(* IEC 61131-3 sources: Caravan/Archiv/12-04-19/Stations/MachineControl/MachineControl/Network/STDPLCInfoPLC, 1 file *)

(* ---- ONE_STDPLCInfoPLC_Table.st ---- *)
#define OBJECTS_CONFIG

#include <.\lsl_st_mt.h>
//Define part of class PLC_Info
#define PLC_INFO_UPDATE_TIME                    250       //Update time in cywork for CPU values
#define PLC_INFO_DEVICE_ID_CPU_REGISTER         16#0F02   //Device ID from wb_cpu_register from  FPGA
#define PLC_INFO_CPU_REGISTER_OFFSET_CPU_TEMP   16#0A     //Offset of wb_cpu_register for CPU Temperature
#define PLC_INFO_CONVERT_TO_1_10_CELSIUS        10        //Multiplier to convert temperature to 1/10°C
#include "..\..\Source\interfaces\lsl_st_pci.h"
#include "..\..\Source\interfaces\lsl_st_syssernum.h"
#include "..\..\Class\PLC_Info\XRegs.h"
#include <.\LoaderItf.h>
#include "..\..\Source\interfaces\lsl_st_sysinfo.h"

FUNCTION GLOBAL TAB ONE_STDPLCInfoPLC
-1$UINT, 0$UINT,
1$UINT, 0$UINT,

7$UDINT,
TO_UDINT(2897291062), "ASCII_BIN", 1$UINT, 20$UINT, 1$UINT,
TO_UDINT(4017734107), "GetOSVersion", 1$UINT, 2$UINT, 1$UINT,
TO_UDINT(2225119864), "MerkerEx", 1$UINT, 22$UINT, 6$UINT,
TO_UDINT(1551372421), "PLC_Info", 1$UINT, 68$UINT, 1$UINT,
TO_UDINT(1850111279), "String", 1$UINT, 10$UINT, 6$UINT,
TO_UDINT(2898603620), "StringInternal", 1$UINT, 82$UINT, 0$UINT,
TO_UDINT(3232495061), "VirtualBaseInit", 1$UINT, 3$UINT, 0$UINT,

_NO_ATTR, TO_UDINT(2882889660), "OSVERSIONPLC",

_NO_ATTR, TO_UDINT(3271492034), "GETOSVERSION_PLC",

1$UINT, TO_UDINT(884148240), "STDPLC_INFOMC1\APPLINAME\MERKEREX0",
1$UINT, TO_UDINT(2112576231), "STDPLC_INFOMC1\CPUBOARD\MERKEREX0",
1$UINT, TO_UDINT(3287353412), "STDPLC_INFOMC1\STRING0\MERKEREX0",
1$UINT, TO_UDINT(41932676), "STDPLC_INFOMC1\STRING1\MERKEREX0",
1$UINT, TO_UDINT(2235530159), "STDPLC_INFOMC1\SYSINFO\MERKEREX0",
1$UINT, TO_UDINT(3997641336), "STRINGOSVERSION_PLC\MERKEREX0",

_NO_ATTR, TO_UDINT(3849002512), "STDPLC_INFOMC1",

1$UINT, TO_UDINT(75928146), "STDPLC_INFOMC1\APPLINAME",
1$UINT, TO_UDINT(3372416669), "STDPLC_INFOMC1\CPUBOARD",
1$UINT, TO_UDINT(1828594461), "STDPLC_INFOMC1\STRING0",
1$UINT, TO_UDINT(469308299), "STDPLC_INFOMC1\STRING1",
1$UINT, TO_UDINT(882984095), "STDPLC_INFOMC1\SYSINFO",
_NO_ATTR, TO_UDINT(3965193377), "STRINGOSVERSION_PLC",

//Internal connections
0$UDINT,
11$UDINT,
TO_UDINT(8), "String0", TO_UDINT(11),
TO_UDINT(8), "String1", TO_UDINT(12),
TO_UDINT(8), "AppliName", TO_UDINT(9),
TO_UDINT(8), "CPUBoard", TO_UDINT(10),
TO_UDINT(8), "SysInfo", TO_UDINT(13),
TO_UDINT(9), "MerkerEx0", TO_UDINT(2),
TO_UDINT(10), "MerkerEx0", TO_UDINT(3),
TO_UDINT(11), "MerkerEx0", TO_UDINT(4),
TO_UDINT(12), "MerkerEx0", TO_UDINT(5),
TO_UDINT(13), "MerkerEx0", TO_UDINT(6),
TO_UDINT(14), "MerkerEx0", TO_UDINT(7),
0$UDINT,
8$UDINT,
TO_UDINT(1), "cOSVersion", TO_UDINT(14), "Data",
TO_UDINT(1), "cAsciiBin", TO_UDINT(0), "Obj_channel",
TO_UDINT(9), "DataBuffer", TO_UDINT(2), "m_udLength",
TO_UDINT(10), "DataBuffer", TO_UDINT(3), "m_udLength",
TO_UDINT(11), "DataBuffer", TO_UDINT(4), "m_udLength",
TO_UDINT(12), "DataBuffer", TO_UDINT(5), "m_udLength",
TO_UDINT(13), "DataBuffer", TO_UDINT(6), "m_udLength",
TO_UDINT(14), "DataBuffer", TO_UDINT(7), "m_udLength",

//Initialization values
0$UDINT,
10$UDINT,
TO_UDINT(2), "ThreadSafe", TO_UDINT(0),//|STDPLCInfoPLC.AppliName\STDPLC_InfoMC1\MerkerEx0.ThreadSafe;
TO_UDINT(3), "ThreadSafe", TO_UDINT(0),//|STDPLCInfoPLC.CPUBoard\STDPLC_InfoMC1\MerkerEx0.ThreadSafe;
TO_UDINT(4), "ThreadSafe", TO_UDINT(0),//|STDPLCInfoPLC.String0\STDPLC_InfoMC1\MerkerEx0.ThreadSafe;
TO_UDINT(5), "ThreadSafe", TO_UDINT(0),//|STDPLCInfoPLC.String1\STDPLC_InfoMC1\MerkerEx0.ThreadSafe;
TO_UDINT(6), "ThreadSafe", TO_UDINT(0),//|STDPLCInfoPLC.SysInfo\STDPLC_InfoMC1\MerkerEx0.ThreadSafe;
TO_UDINT(9), "SingleRealloc", TO_UDINT(1),//|STDPLCInfoPLC.STDPLC_InfoMC1\AppliName.SingleRealloc;
TO_UDINT(10), "SingleRealloc", TO_UDINT(1),//|STDPLCInfoPLC.STDPLC_InfoMC1\CPUBoard.SingleRealloc;
TO_UDINT(11), "SingleRealloc", TO_UDINT(1),//|STDPLCInfoPLC.STDPLC_InfoMC1\String0.SingleRealloc;
TO_UDINT(12), "SingleRealloc", TO_UDINT(1),//|STDPLCInfoPLC.STDPLC_InfoMC1\String1.SingleRealloc;
TO_UDINT(13), "SingleRealloc", TO_UDINT(1),//|STDPLCInfoPLC.STDPLC_InfoMC1\SysInfo.SingleRealloc;

//Symbolic initialization values
0$UDINT,
0$UDINT,

//Initialization of string values
0$UDINT,
0$UDINT,

//Configuration of tasks (RealTime, Cyclic, Background)
0$UDINT,
0$UDINT,

0$UDINT,
0$UDINT,

0$UDINT,
0$UDINT,

//External connections
0$UDINT,
0$UDINT,

//Magic internal connections
0$UDINT,
0$UDINT,

//Configuration of timeslots of tasks (RealTime, Cyclic)
#ifdef __LSLLDR_TIMESLOTS__
0$UDINT,
0$UDINT,

0$UDINT,
0$UDINT,

#endif //__LSLLDR_TIMESLOTS__

//MultiMaster connections
#ifdef __LSLLDR_MULTIMASTER__
0$UDINT,
0$UDINT,
#endif //__LSLLDR_MULTIMASTER__

//Configuration for task ID (RealTime, CyclicTime)
#ifdef __LSLLDR_TASKID__
"\\\\TASKS2  "
0$UDINT,
0$UDINT,

0$UDINT,
0$UDINT,

0$UDINT,
0$UDINT,

#endif //__LSLLDR_TASKID__

END_FUNCTION
